(* IEC 61131-3 sources: PLC-Static-Analysis/modules/plc-rules/src/test/resources/PLCA-L007, 2 files *)

(* ---- compliant.st ---- *)
PROGRAM P_L007ok
VAR
    n : INT;
    m : INT;
    r : REAL;
    b : BOOL;
    c : BOOL;
    q : BOOL;
END_VAR
VAR CONSTANT
    cOn : BOOL := TRUE;
END_VAR
q := r = r;
q := n > 5 OR m <= 5;
q := cOn OR NOT cOn;
q := b OR NOT c;
END_PROGRAM

(* ---- noncompliant.st ---- *)
PROGRAM P_L007
VAR
    n : INT;
    m : INT;
    r : REAL;
    b : BOOL;
    c : BOOL;
    q : BOOL;
END_VAR
IF n > 5 OR n <= 5 THEN // PLCA-L007
    q := TRUE;
END_IF
q := b OR c OR NOT b; // PLCA-L007
q := n = n; // PLCA-L007
q := NOT (b AND NOT b); // PLCA-L007
END_PROGRAM
